(* Logix 5000 project; controller TFF vendor 1 type 14 code 107 rev 33.11; software revision 33.04; part 31 of 38 *)
(* tags used below, declared in another part *)
   Config : Configuration;   // Index Array used in configuration routines
   TIME : DINT[2];
   AC008 : ALIAS FOR DigitalOutput[7];
   AlarmControl : AlarmControl;   // Alarm Control
   ALM002 : ALIAS FOR DigitalOutput[17];
   AnalogOutput : AnalogOutput[25];   // Analog Output Array
   AnalogPoint : AnalogInput[50];   // Analog Input Array
   CCPSystem : CCPSystem;   // CCP System Data
   ChartMark : ChartMark;   // Chart Mark
   Concentration : Concentration;
   CPU_Scanning : BOOL;   // System Scanning Flag
   Diafiltration : Diafiltration;
   DigitalPoint : DigitalPoint[150];   // Digital Point Array
   Drive : Drive[11];   // Drives Array
   FirstScanComplete : BOOL;   // First Scan Complete Flag
   FlowPath : FlowPath[64];   // Flow Path Array
   Gateway : Gateway;   // Gateway Control
   MIX101DF : ALIAS FOR DigitalPoint[28];
   Mixer : Mixer;   // Mixer config. structure
   Operation : Operation[6,251];   // Operation Table
   Options : Options;   // Options List
   Phase0 : ALIAS FOR Phase[0];   // Phase 0
   Phase0_Totalizer_Feed : ALIAS FOR PhaseTotalizer[0];   // Phase 0 Total Feed
   Phase0_Totalizer_Filtrate : ALIAS FOR PhaseTotalizer[6];   // Phase 0 Total Filtrate
   Phase0_Totalizer_Transfer : ALIAS FOR PhaseTotalizer[12];   // Phase 0 Total Transfer
   PipeAnimation : PipeAnimation;   // HMI Pipe Animation Array
   PISL601 : ALIAS FOR DigitalPoint[0];
   PLCFault : FaultRecordType;   // PLC Major Fault Record
   POWERON : ALIAS FOR DigitalOutput[1];
   PTA001 : ALIAS FOR DigitalOutput[21];
   PTA101 : ALIAS FOR DigitalOutput[22];
   PTA201 : ALIAS FOR DigitalOutput[23];
   PTA401 : ALIAS FOR DigitalOutput[24];
   PTA601 : ALIAS FOR DigitalOutput[26];
   PumpRunStatus : DINT;   // Pumps Run Status (1 = At least one pump running , 0 = no pump running)
   Rack_ACT350_WI101_200L : IO_Station;   // Status of ACT350 200L
   Rack_ACT350_WI101_500L : IO_Station;   // Status of ACT350 500L
   SIC001 : ALIAS FOR Drive[1];
   SIC001_AO : ALIAS FOR AnalogOutput[0];
   SIC002 : ALIAS FOR Drive[2];
   SIC002_AO : ALIAS FOR AnalogOutput[1];
   SIC004 : ALIAS FOR Drive[3];
   SysControl : SysControl;   // General system status and command
   Tank : TankManagement;   // Tank Management
   TimerControl : TimerControl;   // Timer Control
   Timers : Timers[22];   // Timer Array
   TNK101 : ALIAS FOR DigitalOutput[18];
   TNK102 : ALIAS FOR DigitalOutput[19];
   TNK103 : ALIAS FOR DigitalOutput[27];
   Totalizer : Totalizers[20];   // Totalizers Array
   UserAlarm : UserAlarm;   // User Alarm (used in CCP Recipe)
   UserCr1 : ALIAS FOR DigitalPoint[65];
   UserCr2 : ALIAS FOR DigitalPoint[67];
   UserNCr1 : ALIAS FOR DigitalPoint[64];
   UserNCr2 : ALIAS FOR DigitalPoint[66];
   UserTime : ALIAS FOR Timers[18];   // User time
   UserTotalizerManagement : UserTotalizerManagement;   // User Totalizer management
   Valve : Valve[100];   // Valve Array
   WI101 : ALIAS FOR AnalogPoint[15];
   YA10 : ALIAS FOR DigitalPoint[59];
   YA41 : ALIAS FOR DigitalPoint[73];
(* Process, continued *)

ROUTINE InputProcessing   (* ladder *)
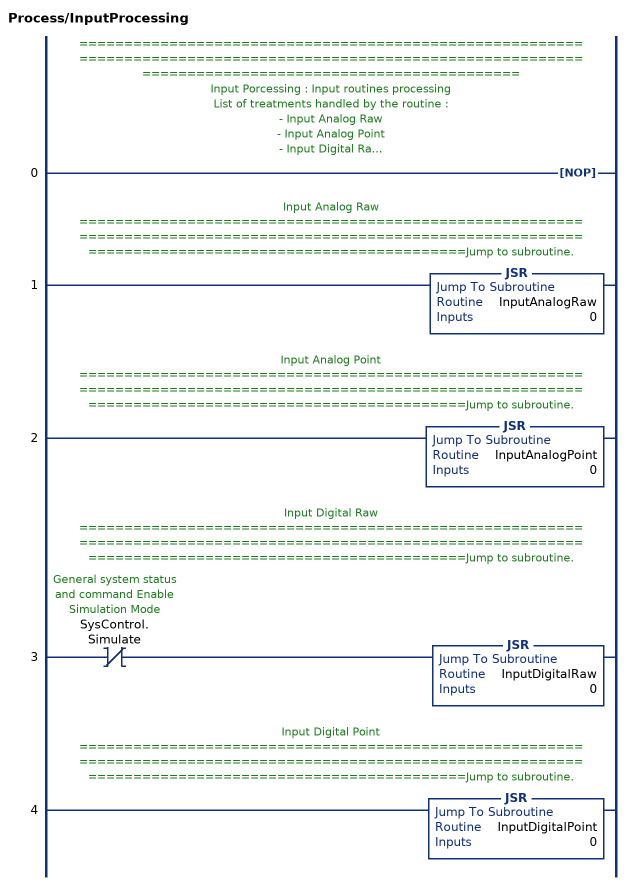
   // ==========================================================================================================================================================
   //                                                                                                                      Input Porcessing : Input routines processing
   //                                                     List of treatments handled by the routine :
   //                                                          - Input Analog Raw
   //                                                          - Input Analog Point
   //                                                          - Input Digital Raw
   //                                                          - Input Digital Point
   //                                                     -----------------------------------------------------------------------------------------------------------------------------------------------------
   //                                                     History
   // 		2019-DEC-24 - Merck - Q. Spindler - Initial version for Candidate Release 1.00.00.00.a
   // ==========================================================================================================================================================
   0: NOP();
   // Input Analog Raw
   // ==========================================================================================================================================================Jump to subroutine.
   1: JSR(InputAnalogRaw,0);
   // Input Analog Point
   // ==========================================================================================================================================================Jump to subroutine.
   2: JSR(InputAnalogPoint,0);
   // Input Digital Raw
   // ==========================================================================================================================================================Jump to subroutine.
   3: XIO(SysControl.Simulate)JSR(InputDigitalRaw,0);
   // Input Digital Point
   // ==========================================================================================================================================================Jump to subroutine.
   4: JSR(InputDigitalPoint,0);
END_ROUTINE

ROUTINE MainRoutine   (* ladder *)
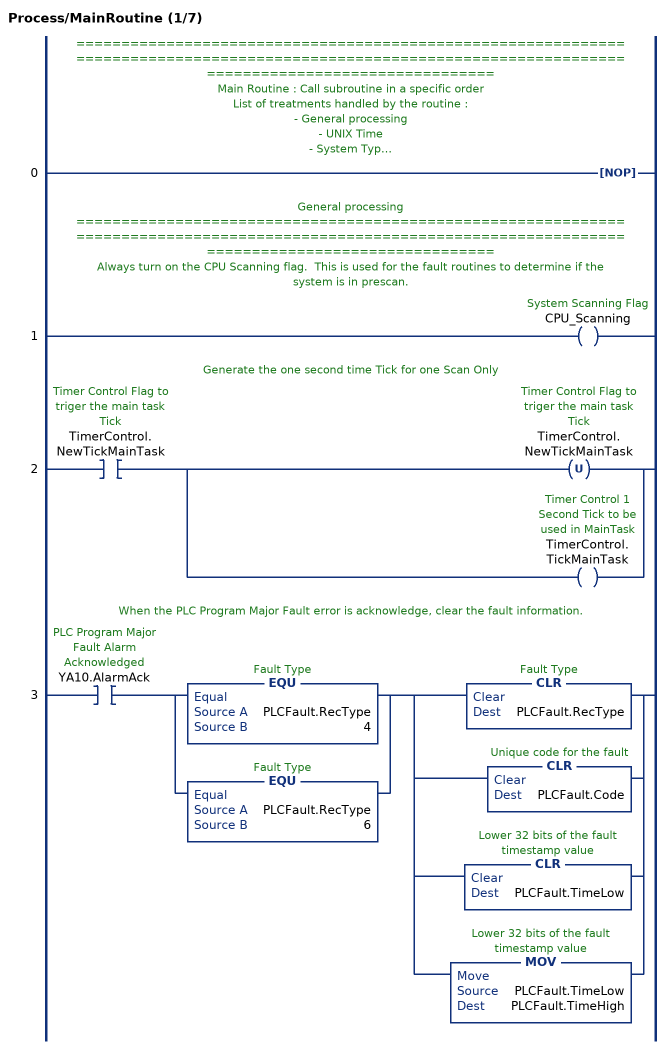
   // ==========================================================================================================================================================
   //                                                                                                            Main Routine : Call subroutine in a specific order
   //                                                     List of treatments handled by the routine :
   //                                                          - General processing
   //                                                          - UNIX Time
   //                                                          - System Type
   //                                                          - Options Configuration
   //                                                         - I/O Station Configuration
   //                                                          - AnalogOutput Configuration
   //                                                          - AnalogPoint Configuration
   //                                                          - DigitalPoint Configuration (real input)
   //                                                          - DigitalPoint Configuration (soft input)
   //                                                          - Valve Configuration
   //                                                          - Drive Configuration
   //                                                          - Control Loop Configuration
   //                                                          - Totalizers Configuration
   //                                                          - Flowpath Configuration
   //                                                          - Reset Configuration
   //                                                          - Station Status
   //                                                          - Derived Data
   //                                                          - Analog and Digital Input Processing
   //                                                         - Modbus Device Processing
   //                                                          - Pump Control
   //                                                          - Loop Control
   //                                                          - Valve Control
   //                                                          - Pipe Animation
   //                                                          - Alarm
   //                                                          - Concentration & Diafiltration
   //                                                          - TankManagement
   //                                                          - Miscellaneous Functions
   //                                                          - Exchange Input and Output
   //                                                          - Analog and Digital Output Processing
   //                                                     - Gateway
   //                                                     -----------------------------------------------------------------------------------------------------------------------------------------------------
   //                                                     History
   // 		2019-DEC-24 - Merck - Q. Spindler - Initial version for Candidate Release 1.00.00.00.a
   // 		2020-APR-06 - Merck - Q. Spindler - Modifications for Candidate Release 1.00.00.00.b
   //                                                 - Add rung to Generate the one second time Tick for one Scan Only
   // ==========================================================================================================================================================
   0: NOP();
   // General processing
   // ==========================================================================================================================================================
   // Always turn on the CPU Scanning flag.  This is used for the fault routines to determine if the system is in prescan.
   1: OTE(CPU_Scanning);
   // Generate the one second time Tick for one Scan Only
   2: XIC(TimerControl.NewTickMainTask)[OTU(TimerControl.NewTickMainTask) ,OTE(TimerControl.TickMainTask) ];
   // When the PLC Program Major Fault error is acknowledge, clear the fault information.
   3: XIC(YA10.AlarmAck)[EQU(PLCFault.RecType,4) ,EQU(PLCFault.RecType,6) ][CLR(PLCFault.RecType) ,CLR(PLCFault.Code) ,CLR(PLCFault.TimeLow) ,MOV(PLCFault.TimeLow,PLCFault.TimeHigh) ];
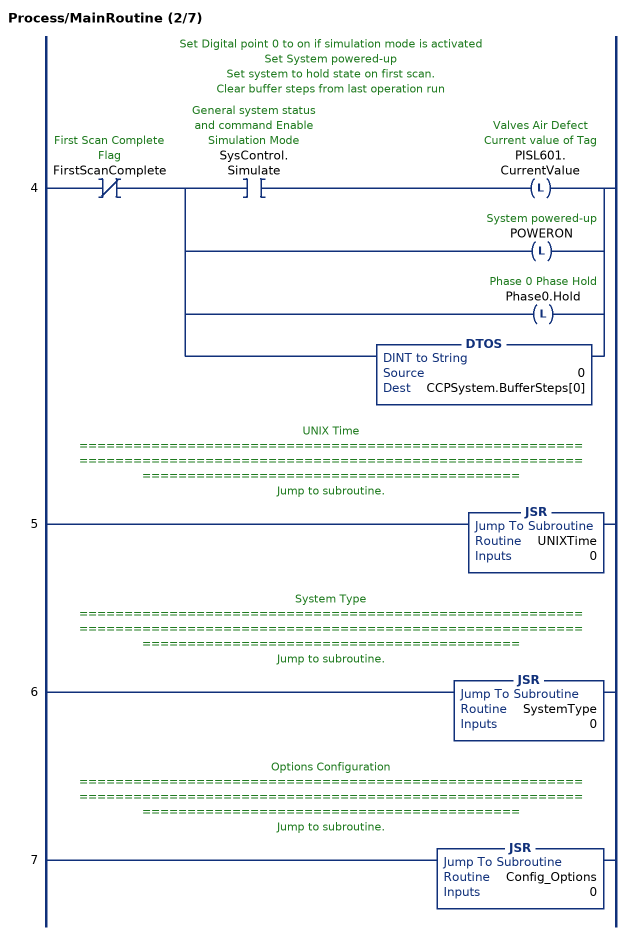
   // Set Digital point 0 to on if simulation mode is activated
   // Set System powered-up
   // Set system to hold state on first scan.
   // Clear buffer steps from last operation run
   4: XIO(FirstScanComplete)[XIC(SysControl.Simulate) OTL(PISL601.CurrentValue) ,OTL(POWERON) ,OTL(Phase0.Hold) ,DTOS(0,CCPSystem.BufferSteps[0]) ];
   // UNIX Time
   // ==========================================================================================================================================================
   // Jump to subroutine.
   5: JSR(UNIXTime,0);
   // System Type
   // ==========================================================================================================================================================
   // Jump to subroutine.
   6: JSR(SystemType,0);
   // Options Configuration
   // ==========================================================================================================================================================
   // Jump to subroutine.
   7: JSR(Config_Options,0);
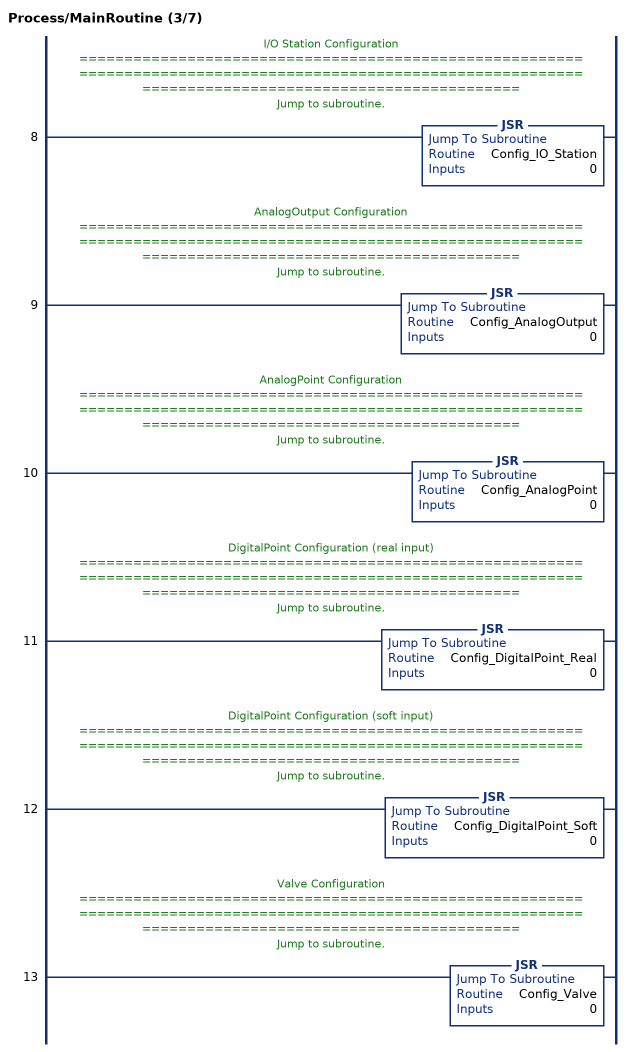
   // I/O Station Configuration
   // ==========================================================================================================================================================
   // Jump to subroutine.
   8: JSR(Config_IO_Station,0);
   // AnalogOutput Configuration
   // ==========================================================================================================================================================
   // Jump to subroutine.
   9: JSR(Config_AnalogOutput,0);
   // AnalogPoint Configuration
   // ==========================================================================================================================================================
   // Jump to subroutine.
   10: JSR(Config_AnalogPoint,0);
   // DigitalPoint Configuration (real input)
   // ==========================================================================================================================================================
   // Jump to subroutine.
   11: JSR(Config_DigitalPoint_Real,0);
   // DigitalPoint Configuration (soft input)
   // ==========================================================================================================================================================
   // Jump to subroutine.
   12: JSR(Config_DigitalPoint_Soft,0);
   // Valve Configuration
   // ==========================================================================================================================================================
   // Jump to subroutine.
   13: JSR(Config_Valve,0);
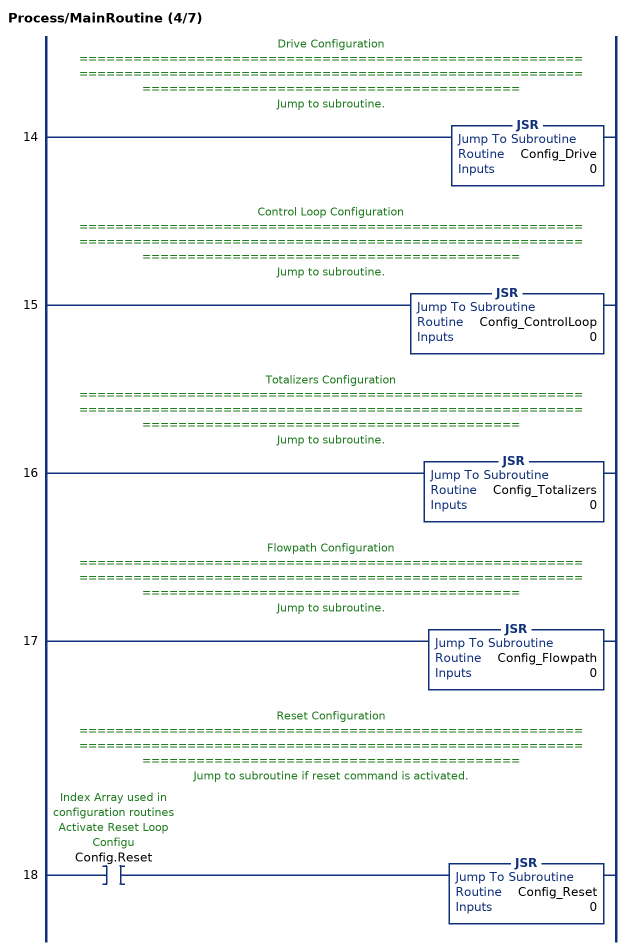
   // Drive Configuration
   // ==========================================================================================================================================================
   // Jump to subroutine.
   14: JSR(Config_Drive,0);
   // Control Loop Configuration
   // ==========================================================================================================================================================
   // Jump to subroutine.
   15: JSR(Config_ControlLoop,0);
   // Totalizers Configuration
   // ==========================================================================================================================================================
   // Jump to subroutine.
   16: JSR(Config_Totalizers,0);
   // Flowpath Configuration
   // ==========================================================================================================================================================
   // Jump to subroutine.
   17: JSR(Config_Flowpath,0);
   // Reset Configuration
   // ==========================================================================================================================================================
   // Jump to subroutine if reset command is activated.
   18: XIC(Config.Reset)JSR(Config_Reset,0);
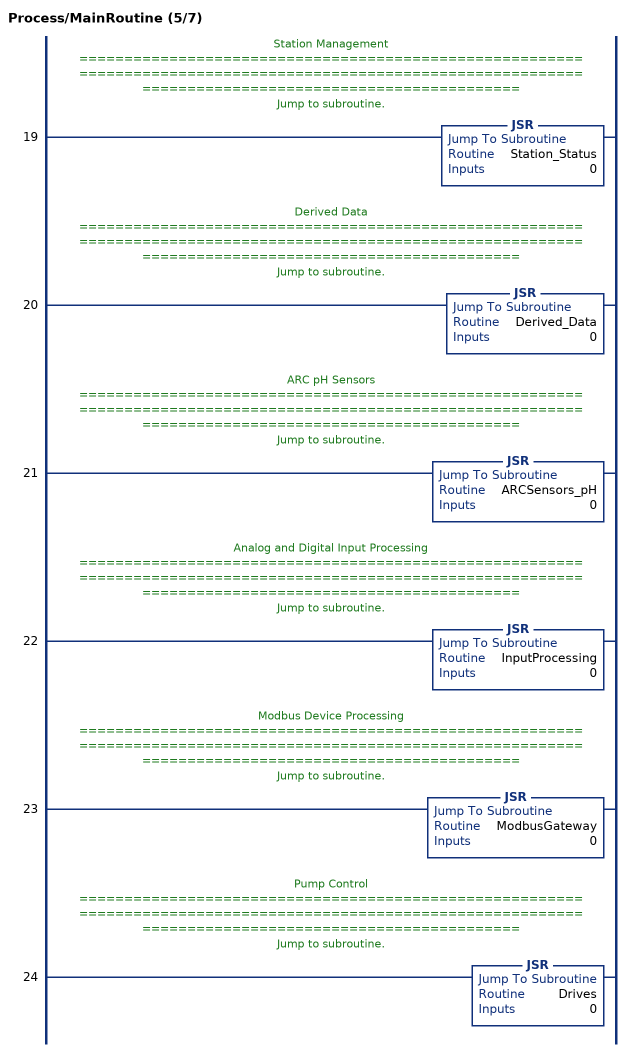
   // Station Management
   // ==========================================================================================================================================================
   // Jump to subroutine.
   19: JSR(Station_Status,0);
   // Derived Data
   // ==========================================================================================================================================================
   // Jump to subroutine.
   20: JSR(Derived_Data,0);
   // ARC pH Sensors
   // ==========================================================================================================================================================
   // Jump to subroutine.
   21: JSR(ARCSensors_pH,0);
   // Analog and Digital Input Processing
   // ==========================================================================================================================================================
   // Jump to subroutine.
   22: JSR(InputProcessing,0);
   // Modbus Device Processing
   // ==========================================================================================================================================================
   // Jump to subroutine.
   23: JSR(ModbusGateway,0);
   // Pump Control
   // ==========================================================================================================================================================
   // Jump to subroutine.
   24: JSR(Drives,0);
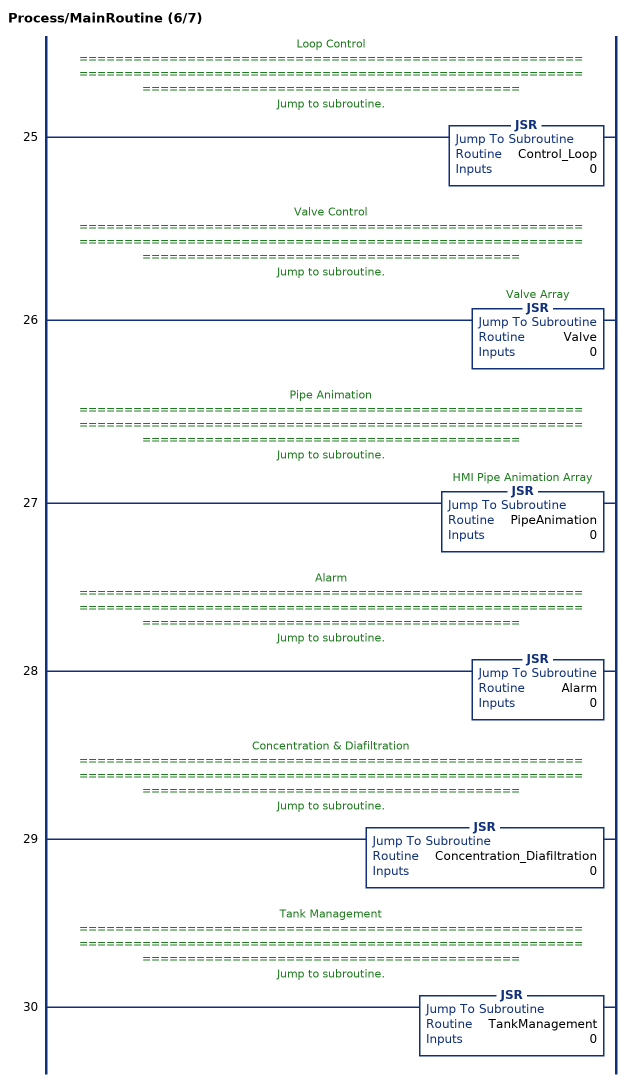
   // Loop Control
   // ==========================================================================================================================================================
   // Jump to subroutine.
   25: JSR(Control_Loop,0);
   // Valve Control
   // ==========================================================================================================================================================
   // Jump to subroutine.
   26: JSR(Valve,0);
   // Pipe Animation
   // ==========================================================================================================================================================
   // Jump to subroutine.
   27: JSR(PipeAnimation,0);
   // Alarm
   // ==========================================================================================================================================================
   // Jump to subroutine.
   28: JSR(Alarm,0);
   // Concentration & Diafiltration
   // ==========================================================================================================================================================
   // Jump to subroutine.
   29: JSR(Concentration_Diafiltration,0);
   // Tank Management
   // ==========================================================================================================================================================
   // Jump to subroutine.
   30: JSR(TankManagement,0);
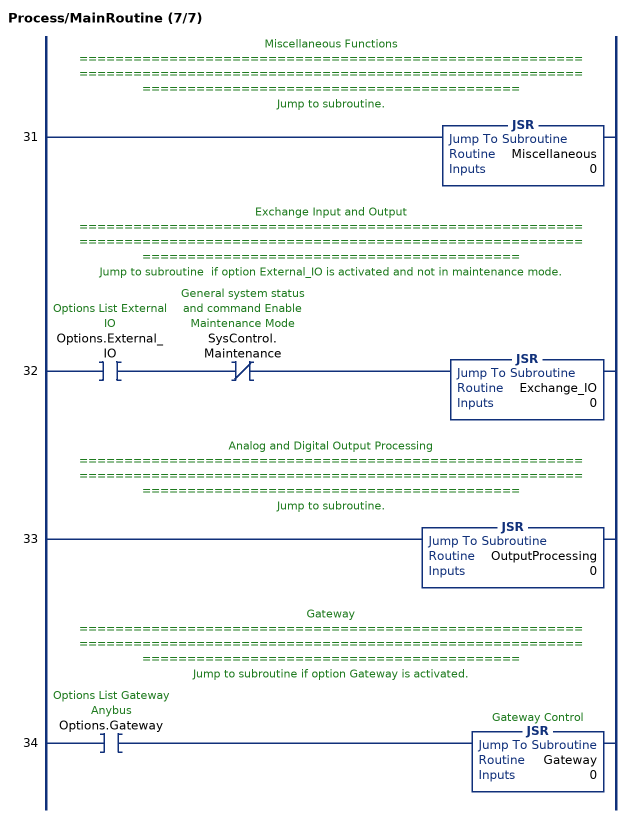
   // Miscellaneous Functions
   // ==========================================================================================================================================================
   // Jump to subroutine.
   31: JSR(Miscellaneous,0);
   // Exchange Input and Output
   // ==========================================================================================================================================================
   // Jump to subroutine  if option External_IO is activated and not in maintenance mode.
   32: XIC(Options.External_IO)XIO(SysControl.Maintenance)JSR(Exchange_IO,0);
   // Analog and Digital Output Processing
   // ==========================================================================================================================================================
   // Jump to subroutine.
   33: JSR(OutputProcessing,0);
   // Gateway
   // ==========================================================================================================================================================
   // Jump to subroutine if option Gateway is activated.
   34: XIC(Options.Gateway)JSR(Gateway,0);
END_ROUTINE

ROUTINE Miscellaneous   (* ladder *)
// Miscellaneous Routine
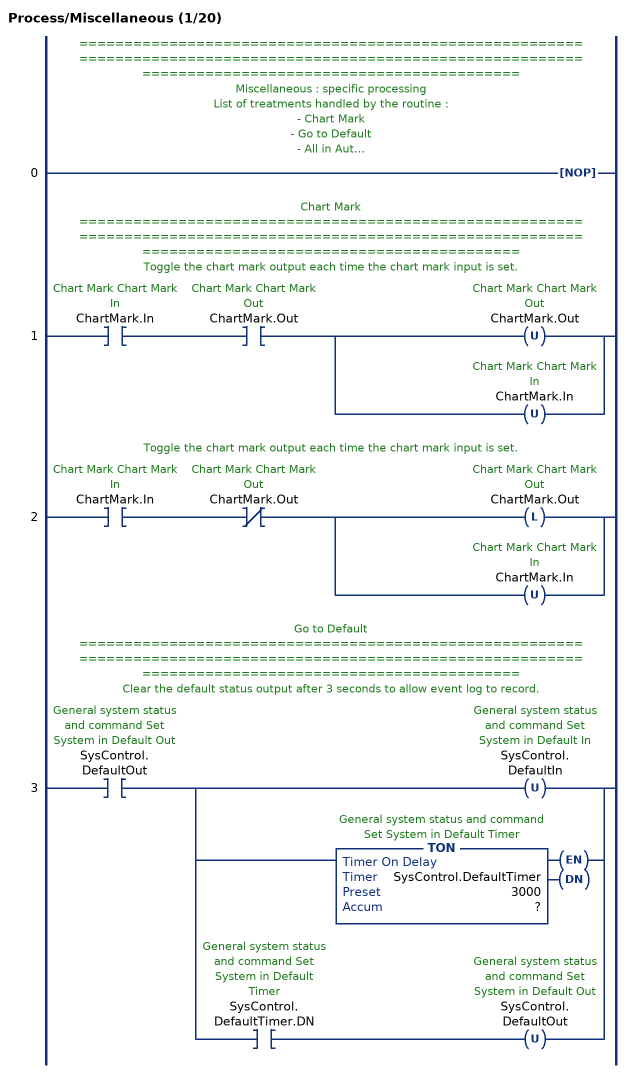
   // ==========================================================================================================================================================
   //                                                                                                                                 Miscellaneous : specific processing
   //                                                     List of treatments handled by the routine :
   //                                                          - Chart Mark
   //                                                          - Go to Default
   //                                                          - All in Auto
   //                                                          - Input Digital Point
   //                                                          - Enable All Alarms
   //                                                          - Disable All Alarms
   //                                                          - Enable all Analog signal alarms
   //                                                          - Disable all Analog signal alarms
   //                                                          - User totalizer management
   //                                                          - Pump Status calculation
   //                                                          - User Alarm (used in recipe only)
   //                                                          - Default Status
   //                                                          - Save \ Restore parameters conditions
   //                                                          - Mixer Reset Alarm Command
   //                                                          - ACT350 Configurations
   //                                                          - UV Baseline Zero Command Logic
   //                                                          - Weight Tare Command Logic
   //                                                         - Pressure Tare Command Logic
   //                                                       - Membrane Status
   //                                                     - C8000 Powerup
   //                                                    - Bag Inflate
   //                                                     - TFF80 Dual Pump managment
   //                                                     - Operating Time Exceeded (YA41)
   //                                                     -----------------------------------------------------------------------------------------------------------------------------------------------------
   //                                                     History
   // 		2019-DEC-24 - Merck - Q. Spindler - Initial version for Candidate Release 1.00.00.00.a
   //                                2020-MAR-25 - Merck - Q. Spindler - Modifications for Candidate Release 1.00.00.00.b
   //                                                                                                            - TFF80 Dual Pump managment, SIC001_AO was copied to SIC002_AO instead of the other way around.
   // - Add WI101 Weight Zero Output
   //                                2021-NOV-22 - Merck - Q. Spindler - Modifications for Candidate Release 1.01.00.00.a
   //   - Add Operating Time Exceeded (YA41)
   // - Add Transfer totalisers (for user totalizer)
   //                                2022-SEP-21 - Actemium - J. Jaekel - Modifications for Candidate Release 1.01.00.01.a
   // - Disable the inflate output cmd when the system is hold
   // ==========================================================================================================================================================
   0: NOP();
   // Chart Mark
   // ==========================================================================================================================================================
   // Toggle the chart mark output each time the chart mark input is set.
   1: XIC(ChartMark.In)XIC(ChartMark.Out)[OTU(ChartMark.Out) ,OTU(ChartMark.In) ];
   // Toggle the chart mark output each time the chart mark input is set.
   2: XIC(ChartMark.In)XIO(ChartMark.Out)[OTL(ChartMark.Out) ,OTU(ChartMark.In) ];
   // Go to Default
   // ==========================================================================================================================================================
   // Clear the default status output after 3 seconds to allow event log to record.
   3: XIC(SysControl.DefaultOut)[OTU(SysControl.DefaultIn) ,TON(SysControl.DefaultTimer,?,?) ,XIC(SysControl.DefaultTimer.DN) OTU(SysControl.DefaultOut) ];
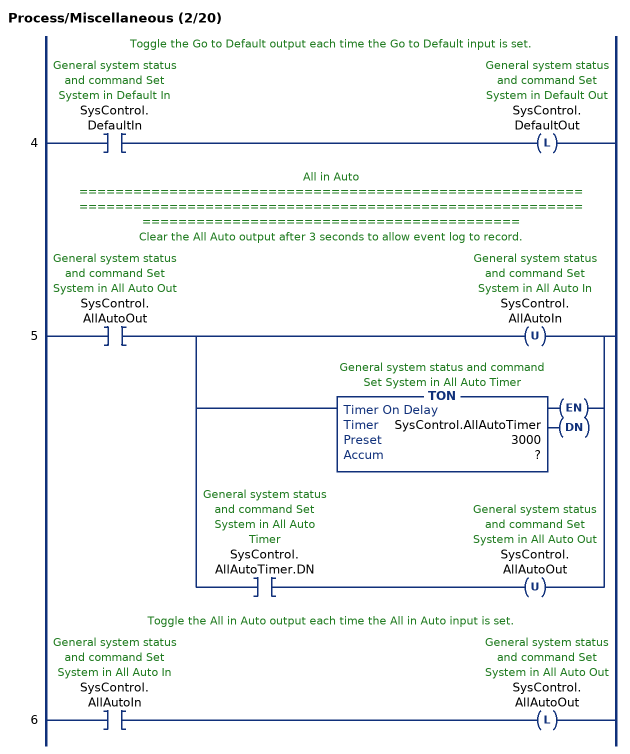
   // Toggle the Go to Default output each time the Go to Default input is set.
   4: XIC(SysControl.DefaultIn)OTL(SysControl.DefaultOut);
   // All in Auto
   // ==========================================================================================================================================================
   // Clear the All Auto output after 3 seconds to allow event log to record.
   5: XIC(SysControl.AllAutoOut)[OTU(SysControl.AllAutoIn) ,TON(SysControl.AllAutoTimer,?,?) ,XIC(SysControl.AllAutoTimer.DN) OTU(SysControl.AllAutoOut) ];
   // Toggle the All in Auto output each time the All in Auto input is set.
   6: XIC(SysControl.AllAutoIn)OTL(SysControl.AllAutoOut);
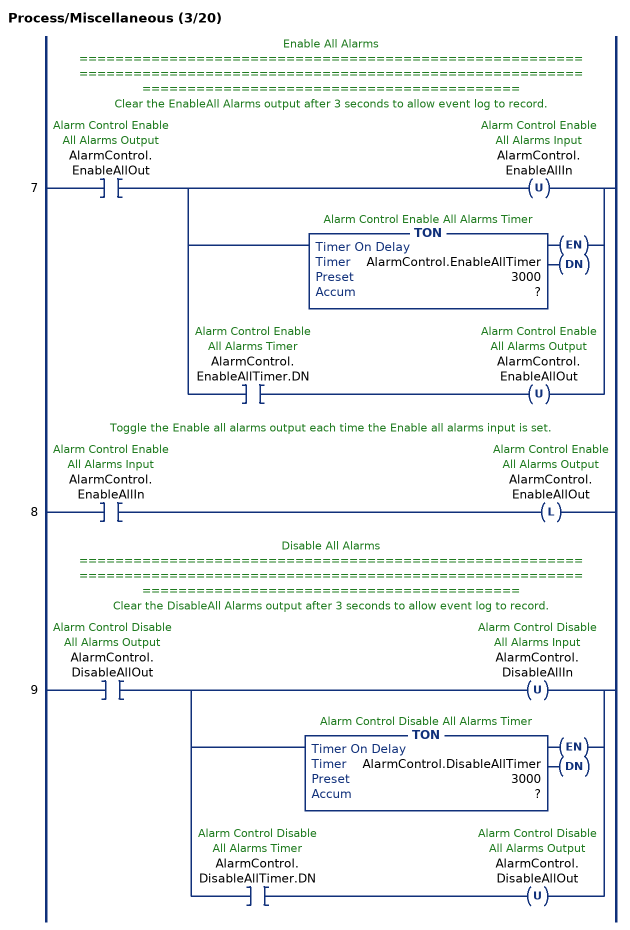
   // Enable All Alarms
   // ==========================================================================================================================================================
   // Clear the EnableAll Alarms output after 3 seconds to allow event log to record.
   7: XIC(AlarmControl.EnableAllOut)[OTU(AlarmControl.EnableAllIn) ,TON(AlarmControl.EnableAllTimer,?,?) ,XIC(AlarmControl.EnableAllTimer.DN) OTU(AlarmControl.EnableAllOut) ];
   // Toggle the Enable all alarms output each time the Enable all alarms input is set.
   8: XIC(AlarmControl.EnableAllIn)OTL(AlarmControl.EnableAllOut);
   // Disable All Alarms
   // ==========================================================================================================================================================
   // Clear the DisableAll Alarms output after 3 seconds to allow event log to record.
   9: XIC(AlarmControl.DisableAllOut)[OTU(AlarmControl.DisableAllIn) ,TON(AlarmControl.DisableAllTimer,?,?) ,XIC(AlarmControl.DisableAllTimer.DN) OTU(AlarmControl.DisableAllOut) ];
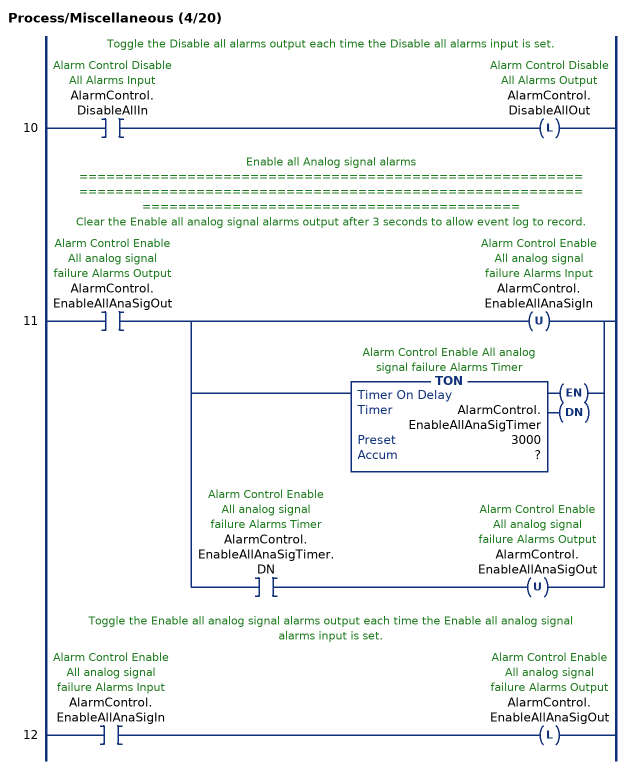
   // Toggle the Disable all alarms output each time the Disable all alarms input is set.
   10: XIC(AlarmControl.DisableAllIn)OTL(AlarmControl.DisableAllOut);
   // Enable all Analog signal alarms
   // ==========================================================================================================================================================
   // Clear the Enable all analog signal alarms output after 3 seconds to allow event log to record.
   11: XIC(AlarmControl.EnableAllAnaSigOut)[OTU(AlarmControl.EnableAllAnaSigIn) ,TON(AlarmControl.EnableAllAnaSigTimer,?,?) ,XIC(AlarmControl.EnableAllAnaSigTimer.DN) OTU(AlarmControl.EnableAllAnaSigOut) ];
   // Toggle the Enable all analog signal alarms output each time the Enable all analog signal alarms input is set.
   12: XIC(AlarmControl.EnableAllAnaSigIn)OTL(AlarmControl.EnableAllAnaSigOut);
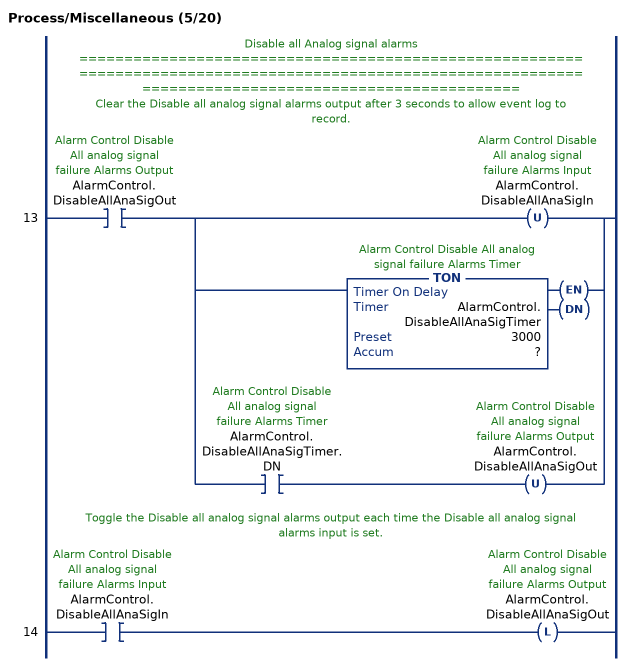
   // Disable all Analog signal alarms
   // ==========================================================================================================================================================
   // Clear the Disable all analog signal alarms output after 3 seconds to allow event log to record.
   13: XIC(AlarmControl.DisableAllAnaSigOut)[OTU(AlarmControl.DisableAllAnaSigIn) ,TON(AlarmControl.DisableAllAnaSigTimer,?,?) ,XIC(AlarmControl.DisableAllAnaSigTimer.DN) OTU(AlarmControl.DisableAllAnaSigOut) ];
   // Toggle the Disable all analog signal alarms output each time the Disable all analog signal alarms input is set.
   14: XIC(AlarmControl.DisableAllAnaSigIn)OTL(AlarmControl.DisableAllAnaSigOut);
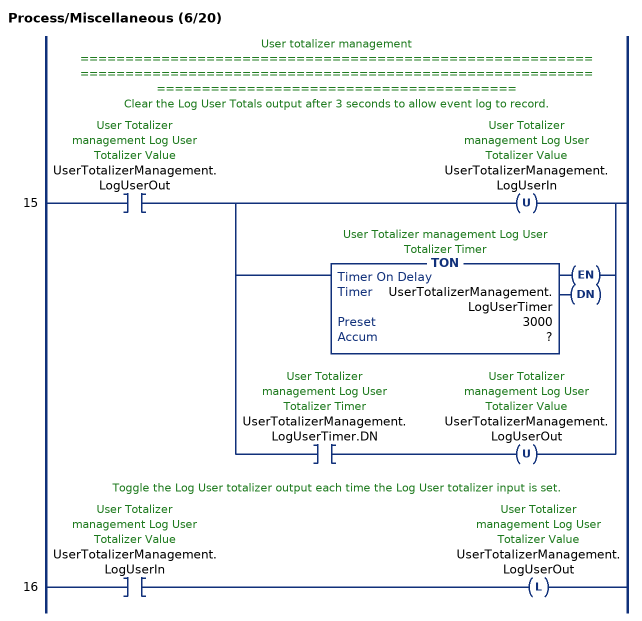
   // User totalizer management
   // ==========================================================================================================================================================
   // Clear the Log User Totals output after 3 seconds to allow event log to record.
   15: XIC(UserTotalizerManagement.LogUserOut)[OTU(UserTotalizerManagement.LogUserIn) ,TON(UserTotalizerManagement.LogUserTimer,?,?) ,XIC(UserTotalizerManagement.LogUserTimer.DN) OTU(UserTotalizerManagement.LogUserOut) ];
   // Toggle the Log User totalizer output each time the Log User totalizer input is set.
   16: XIC(UserTotalizerManagement.LogUserIn)OTL(UserTotalizerManagement.LogUserOut);
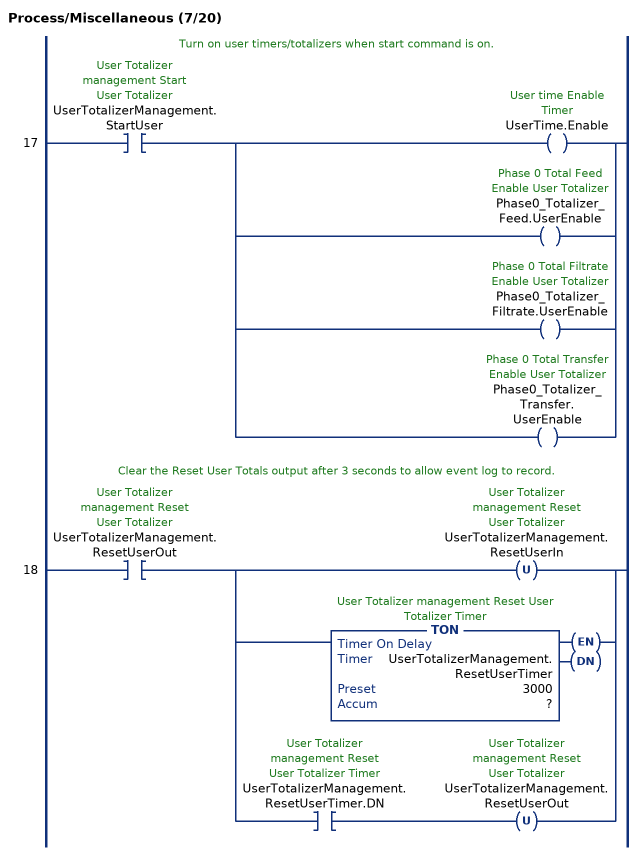
   // Turn on user timers/totalizers when start command is on.
   17: XIC(UserTotalizerManagement.StartUser)[OTE(UserTime.Enable) ,OTE(Phase0_Totalizer_Feed.UserEnable) ,OTE(Phase0_Totalizer_Filtrate.UserEnable) ,OTE(Phase0_Totalizer_Transfer.UserEnable) ];
   // Clear the Reset User Totals output after 3 seconds to allow event log to record.
   18: XIC(UserTotalizerManagement.ResetUserOut)[OTU(UserTotalizerManagement.ResetUserIn) ,TON(UserTotalizerManagement.ResetUserTimer,?,?) ,XIC(UserTotalizerManagement.ResetUserTimer.DN) OTU(UserTotalizerManagement.ResetUserOut) ];
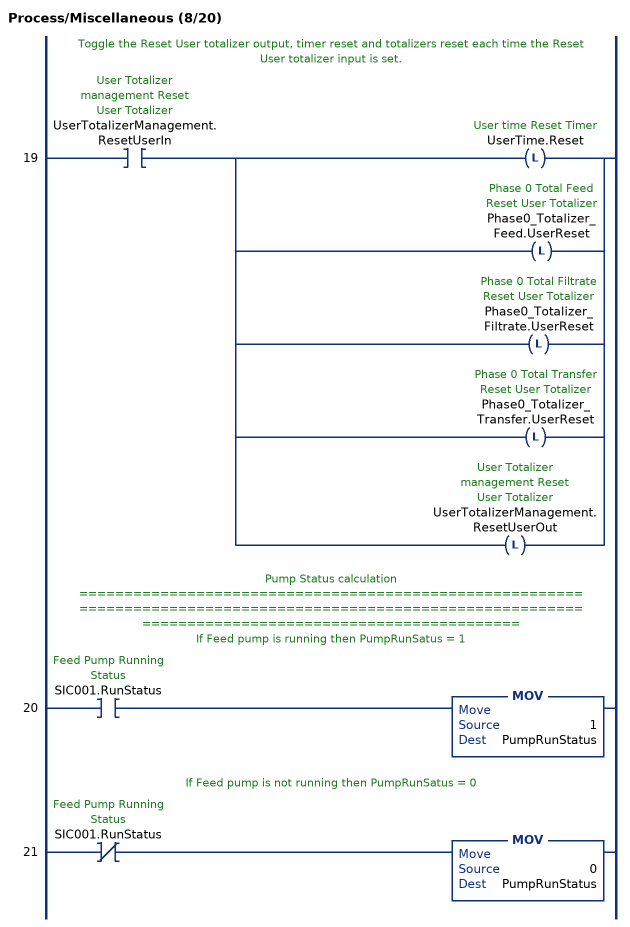
   // Toggle the Reset User totalizer output, timer reset and totalizers reset each time the Reset User totalizer input is set.
   19: XIC(UserTotalizerManagement.ResetUserIn)[OTL(UserTime.Reset) ,OTL(Phase0_Totalizer_Feed.UserReset) ,OTL(Phase0_Totalizer_Filtrate.UserReset) ,OTL(Phase0_Totalizer_Transfer.UserReset) ,OTL(UserTotalizerManagement.ResetUserOut) ];
   // Pump Status calculation
   // ==========================================================================================================================================================
   // If Feed pump is running then PumpRunSatus = 1
   20: XIC(SIC001.RunStatus)MOV(1,PumpRunStatus);
   // If Feed pump is not running then PumpRunSatus = 0
   21: XIO(SIC001.RunStatus)MOV(0,PumpRunStatus);
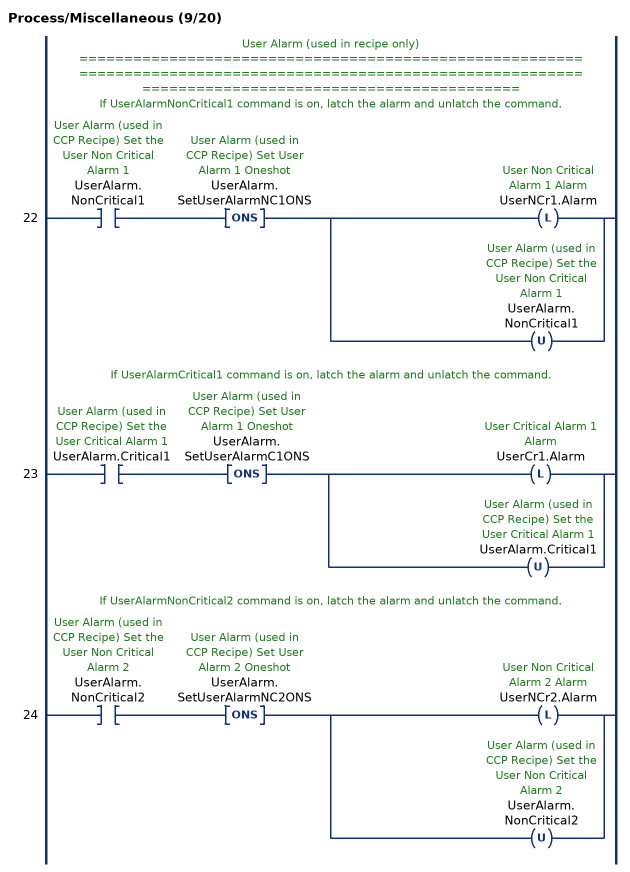
   // User Alarm (used in recipe only)
   // ==========================================================================================================================================================
   // If UserAlarmNonCritical1 command is on, latch the alarm and unlatch the command.
   22: XIC(UserAlarm.NonCritical1)ONS(UserAlarm.SetUserAlarmNC1ONS)[OTL(UserNCr1.Alarm) ,OTU(UserAlarm.NonCritical1) ];
   // If UserAlarmCritical1 command is on, latch the alarm and unlatch the command.
   23: XIC(UserAlarm.Critical1)ONS(UserAlarm.SetUserAlarmC1ONS)[OTL(UserCr1.Alarm) ,OTU(UserAlarm.Critical1) ];
   // If UserAlarmNonCritical2 command is on, latch the alarm and unlatch the command.
   24: XIC(UserAlarm.NonCritical2)ONS(UserAlarm.SetUserAlarmNC2ONS)[OTL(UserNCr2.Alarm) ,OTU(UserAlarm.NonCritical2) ];
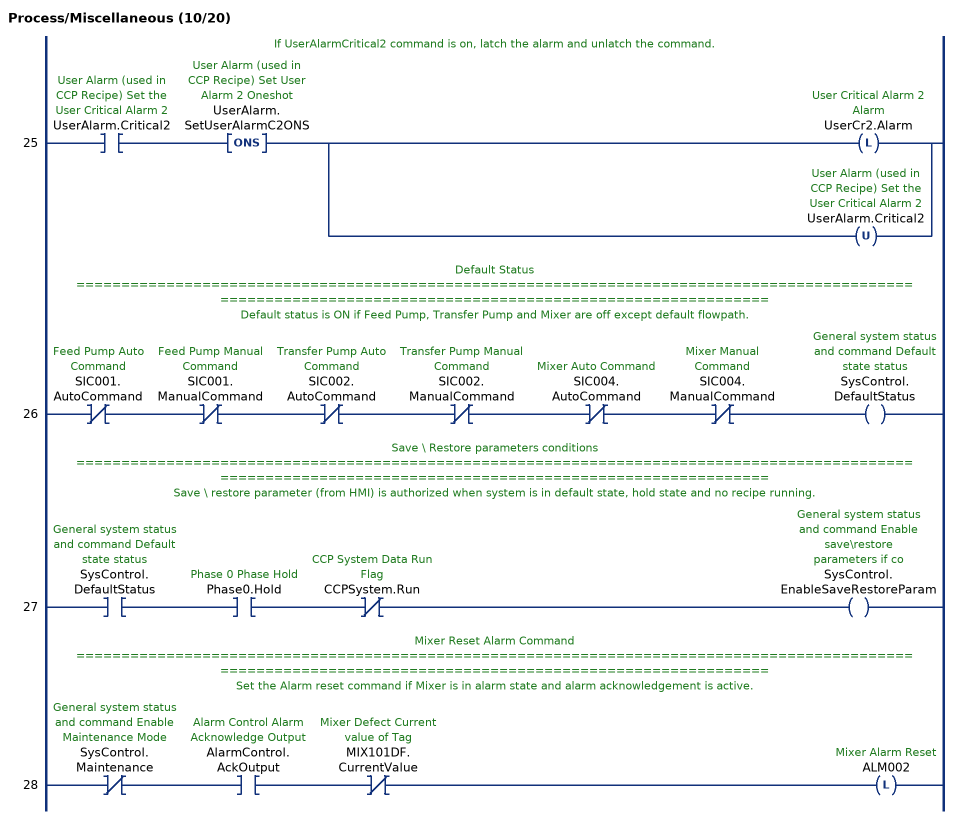
   // If UserAlarmCritical2 command is on, latch the alarm and unlatch the command.
   25: XIC(UserAlarm.Critical2)ONS(UserAlarm.SetUserAlarmC2ONS)[OTL(UserCr2.Alarm) ,OTU(UserAlarm.Critical2) ];
   // Default Status
   // ==========================================================================================================================================================
   // Default status is ON if Feed Pump, Transfer Pump and Mixer are off except default flowpath.
   26: XIO(SIC001.AutoCommand)XIO(SIC001.ManualCommand)XIO(SIC002.AutoCommand)XIO(SIC002.ManualCommand)XIO(SIC004.AutoCommand)XIO(SIC004.ManualCommand)OTE(SysControl.DefaultStatus);
   // Save \ Restore parameters conditions
   // ==========================================================================================================================================================
   // Save \ restore parameter (from HMI) is authorized when system is in default state, hold state and no recipe running.
   27: XIC(SysControl.DefaultStatus)XIC(Phase0.Hold)XIO(CCPSystem.Run)OTE(SysControl.EnableSaveRestoreParam);
   // Mixer Reset Alarm Command
   // ==========================================================================================================================================================
   // Set the Alarm reset command if Mixer is in alarm state and alarm acknowledgement is active.
   28: XIO(SysControl.Maintenance)XIC(AlarmControl.AckOutput)XIO(MIX101DF.CurrentValue)OTL(ALM002);
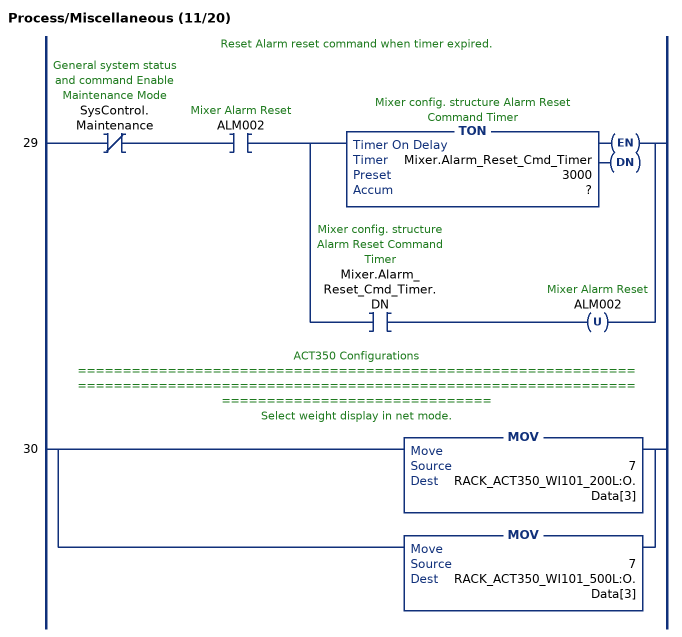
   // Reset Alarm reset command when timer expired.
   29: XIO(SysControl.Maintenance)XIC(ALM002)[TON(Mixer.Alarm_Reset_Cmd_Timer,?,?) ,XIC(Mixer.Alarm_Reset_Cmd_Timer.DN) OTU(ALM002) ];
   // ACT350 Configurations
   // ==========================================================================================================================================================
   // Select weight display in net mode.
   30: [MOV(7,RACK_ACT350_WI101_200L:O.Data[3]) ,MOV(7,RACK_ACT350_WI101_500L:O.Data[3]) ];
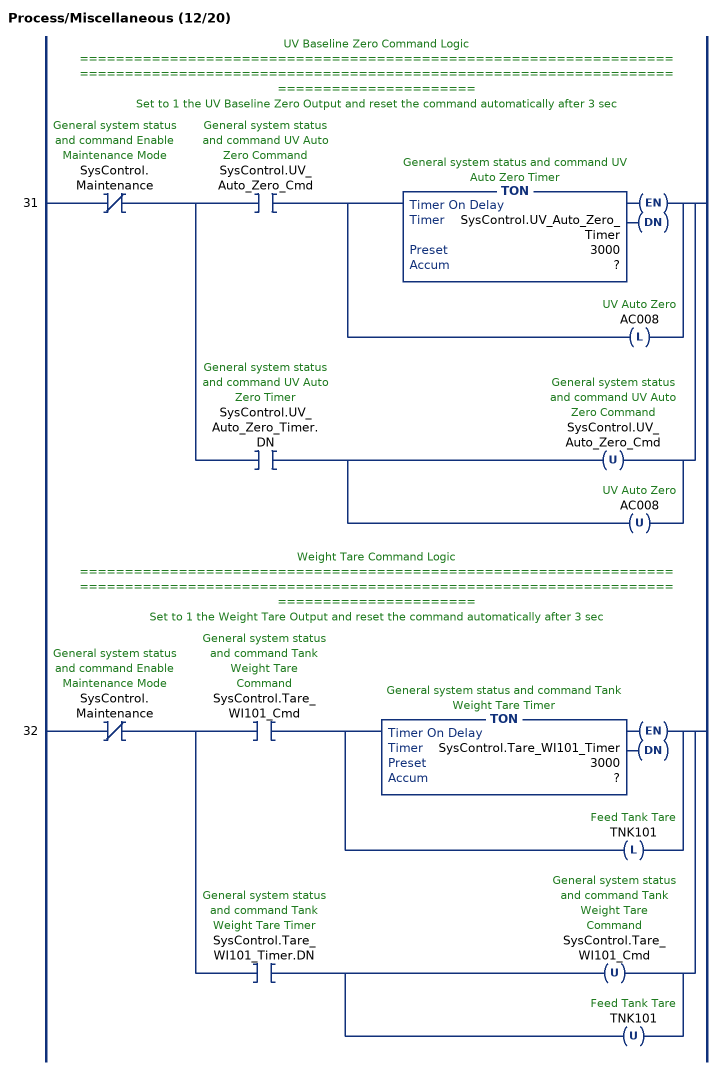
   // UV Baseline Zero Command Logic
   // ==========================================================================================================================================================
   // Set to 1 the UV Baseline Zero Output and reset the command automatically after 3 sec
   31: XIO(SysControl.Maintenance)[XIC(SysControl.UV_Auto_Zero_Cmd) [TON(SysControl.UV_Auto_Zero_Timer,?,?) ,OTL(AC008) ] ,XIC(SysControl.UV_Auto_Zero_Timer.DN) [OTU(SysControl.UV_Auto_Zero_Cmd) ,OTU(AC008) ] ];
   // Weight Tare Command Logic
   // ==========================================================================================================================================================
   // Set to 1 the Weight Tare Output and reset the command automatically after 3 sec
   32: XIO(SysControl.Maintenance)[XIC(SysControl.Tare_WI101_Cmd) [TON(SysControl.Tare_WI101_Timer,?,?) ,OTL(TNK101) ] ,XIC(SysControl.Tare_WI101_Timer.DN) [OTU(SysControl.Tare_WI101_Cmd) ,OTU(TNK101) ] ];
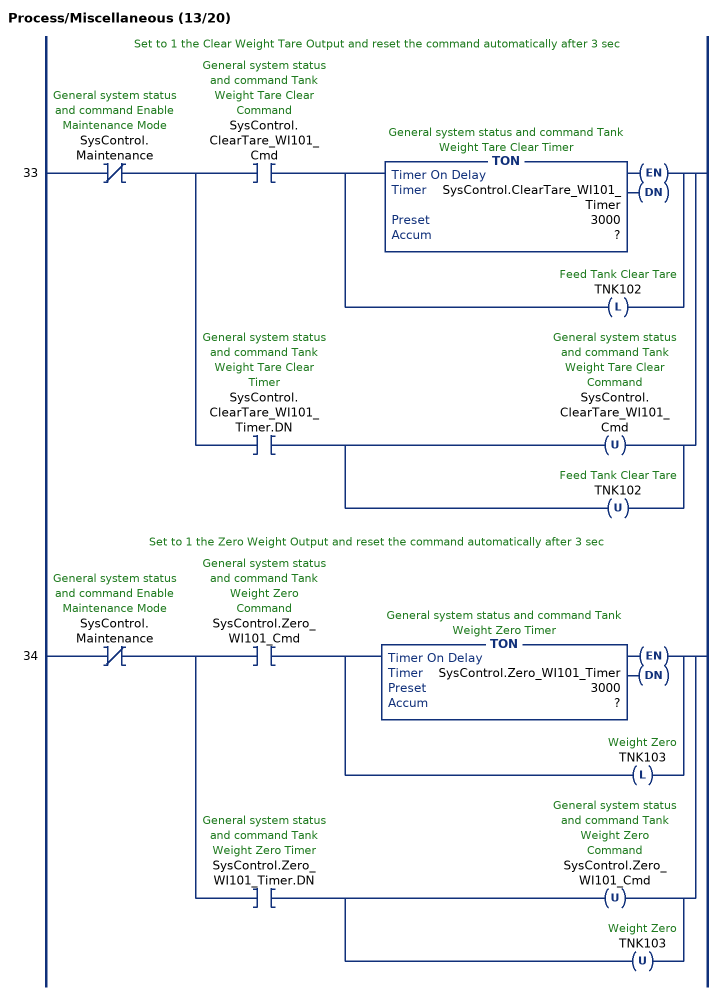
   // Set to 1 the Clear Weight Tare Output and reset the command automatically after 3 sec
   33: XIO(SysControl.Maintenance)[XIC(SysControl.ClearTare_WI101_Cmd) [TON(SysControl.ClearTare_WI101_Timer,?,?) ,OTL(TNK102) ] ,XIC(SysControl.ClearTare_WI101_Timer.DN) [OTU(SysControl.ClearTare_WI101_Cmd) ,OTU(TNK102) ] ];
   // Set to 1 the Zero Weight Output and reset the command automatically after 3 sec
   34: XIO(SysControl.Maintenance)[XIC(SysControl.Zero_WI101_Cmd) [TON(SysControl.Zero_WI101_Timer,?,?) ,OTL(TNK103) ] ,XIC(SysControl.Zero_WI101_Timer.DN) [OTU(SysControl.Zero_WI101_Cmd) ,OTU(TNK103) ] ];
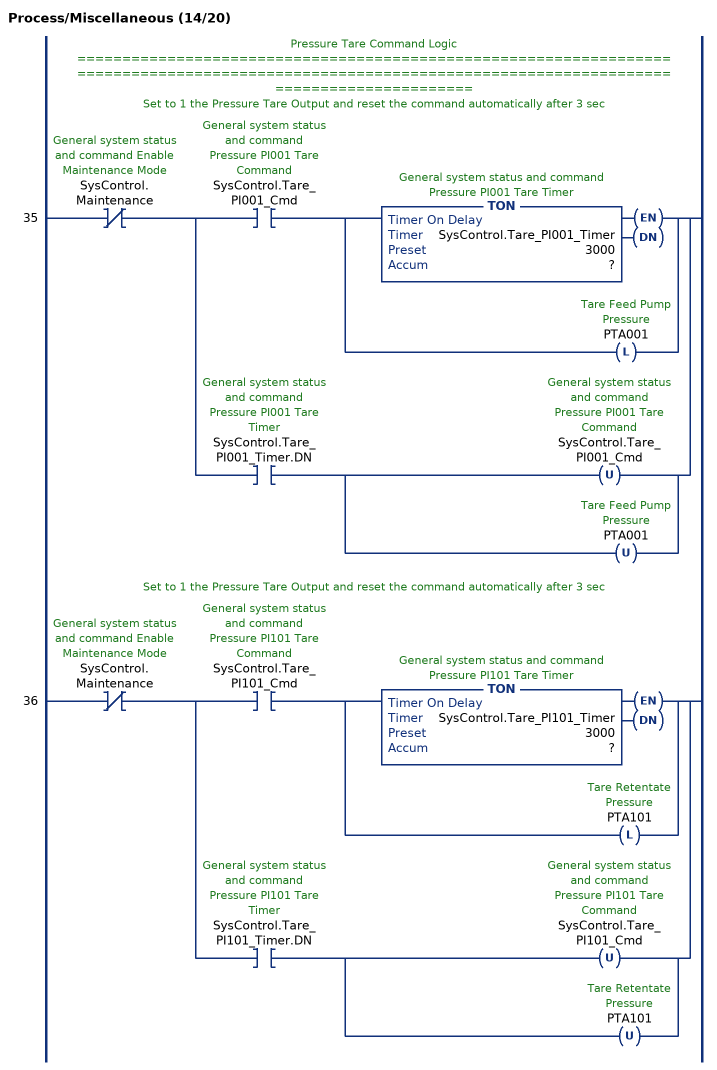
   // Pressure Tare Command Logic
   // ==========================================================================================================================================================
   // Set to 1 the Pressure Tare Output and reset the command automatically after 3 sec
   35: XIO(SysControl.Maintenance)[XIC(SysControl.Tare_PI001_Cmd) [TON(SysControl.Tare_PI001_Timer,?,?) ,OTL(PTA001) ] ,XIC(SysControl.Tare_PI001_Timer.DN) [OTU(SysControl.Tare_PI001_Cmd) ,OTU(PTA001) ] ];
   // Set to 1 the Pressure Tare Output and reset the command automatically after 3 sec
   36: XIO(SysControl.Maintenance)[XIC(SysControl.Tare_PI101_Cmd) [TON(SysControl.Tare_PI101_Timer,?,?) ,OTL(PTA101) ] ,XIC(SysControl.Tare_PI101_Timer.DN) [OTU(SysControl.Tare_PI101_Cmd) ,OTU(PTA101) ] ];
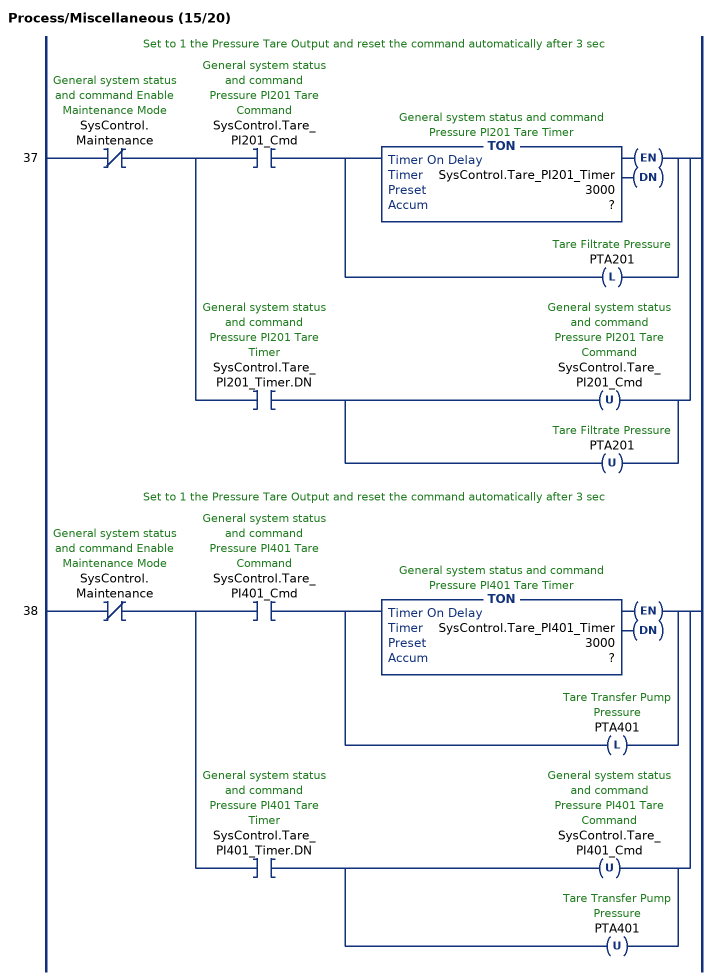
   // Set to 1 the Pressure Tare Output and reset the command automatically after 3 sec
   37: XIO(SysControl.Maintenance)[XIC(SysControl.Tare_PI201_Cmd) [TON(SysControl.Tare_PI201_Timer,?,?) ,OTL(PTA201) ] ,XIC(SysControl.Tare_PI201_Timer.DN) [OTU(SysControl.Tare_PI201_Cmd) ,OTU(PTA201) ] ];
   // Set to 1 the Pressure Tare Output and reset the command automatically after 3 sec
   38: XIO(SysControl.Maintenance)[XIC(SysControl.Tare_PI401_Cmd) [TON(SysControl.Tare_PI401_Timer,?,?) ,OTL(PTA401) ] ,XIC(SysControl.Tare_PI401_Timer.DN) [OTU(SysControl.Tare_PI401_Cmd) ,OTU(PTA401) ] ];
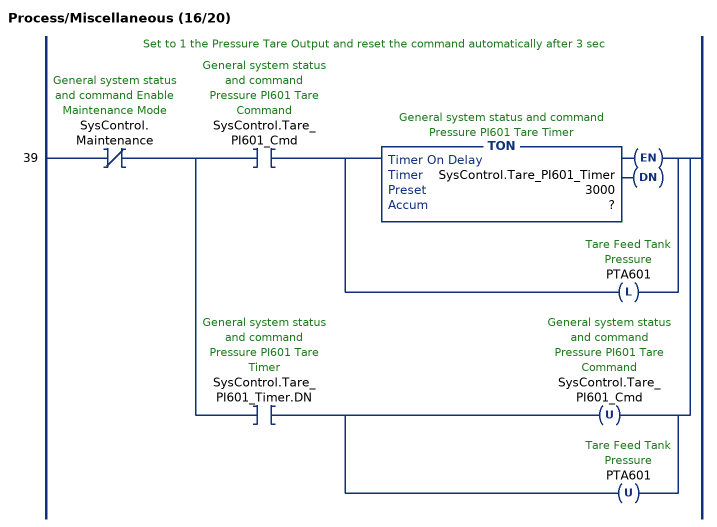
   // Set to 1 the Pressure Tare Output and reset the command automatically after 3 sec
   39: XIO(SysControl.Maintenance)[XIC(SysControl.Tare_PI601_Cmd) [TON(SysControl.Tare_PI601_Timer,?,?) ,OTL(PTA601) ] ,XIC(SysControl.Tare_PI601_Timer.DN) [OTU(SysControl.Tare_PI601_Cmd) ,OTU(PTA601) ] ];
